Fanuc TP program (LS listing): ConfPr.LS

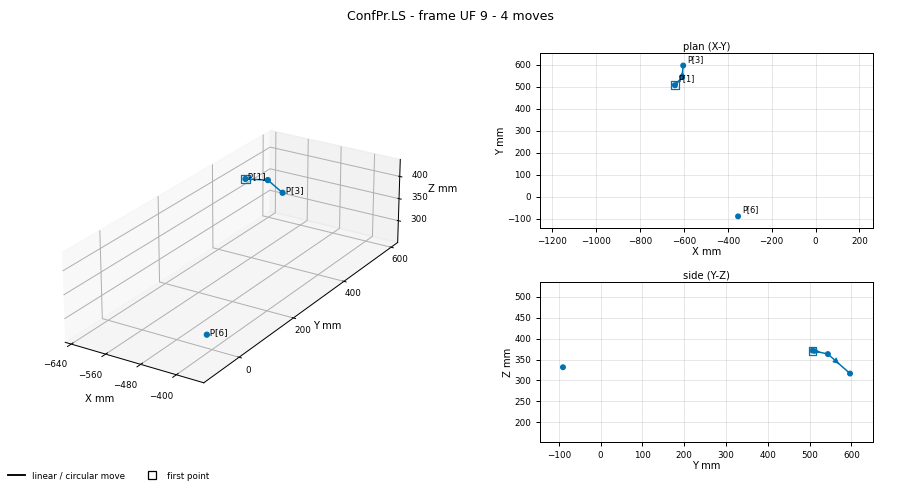
[picture p0: tool path of ConfPr.LS in frame UF 9, 4 of 6 moves have a stored position in this frame; points joined in program order, loops and branches not executed]
/PROG  ConfPr
/ATTR
OWNER		= MNEDITOR;
COMMENT		= "RoboDK sequence";
PROG_SIZE	= 0;
CREATE		= DATE 31-12-14  TIME 12:00:00;
MODIFIED	= DATE 31-12-14  TIME 12:00:00;
FILE_NAME	= ConfPr;
VERSION		= 0;
LINE_COUNT	= 25;
MEMORY_SIZE	= 0;
PROTECT		= READ_WRITE;
TCD:  STACK_SIZE	= 0,
      TASK_PRIORITY	= 50,
      TIME_SLICE	= 0,
      BUSY_LAMP_OFF	= 0,
      ABORT_REQUEST	= 0,
      PAUSE_REQUEST	= 0;
DEFAULT_GROUP	= 1,*,*,*,*;
CONTROL_CODE	= 00000000 00000000;
/MN
   1:  ! Program generated by RoboDK v6.0.7 for Fanuc M-1iA/0.5S on XX ;
   2:  ! /XX/XXXX 18:00:00 ;
   3:  ! Using nominal kinematics. ;
   4:  PR[9,1]=1234.570 ;
   5:  PR[9,2]=-98.765 ;
   6:  PR[9,3]=50.500 ;
   7:  PR[9,4]=0.000 ;
   8:  PR[9,5]=0.000 ;
   9:  PR[9,6]=30.000 ;
  10:  UFRAME[9]=PR[9] ;
  11:  UFRAME_NUM=9 ;
  12:  PR[9,1]=10.000 ;
  13:  PR[9,2]=20.000 ;
  14:  PR[9,3]=150.000 ;
  15:  PR[9,4]=0.000 ;
  16:  PR[9,5]=0.000 ;
  17:  PR[9,6]=0.000 ;
  18:  UTOOL[9]=PR[9] ;
  19:  UTOOL_NUM=9 ;
  20:L P[1] 200mm/sec FINE ;
  21:L P[2] 200mm/sec FINE ;
  22:L P[3] 200mm/sec FINE ;
  23:J P[4] 20% FINE ;
  24:J P[5] 20% FINE ;
  25:C P[6]
       P[7] 200mm/sec FINE ;
/POS
P[1]{
   GP1:
    UF : 9, UT : 9,        CONFIG : 'L, 0, 0, 0',
	X =  -640.584  mm,	Y =   506.980  mm,	Z =   371.534  mm,
	W =  -165.000 deg,	P =    50.000 deg,	R =   150.000 deg
};
P[2]{
   GP1:
    UF : 9, UT : 9,        CONFIG : 'L, 0, 0, 1',
	X =  -607.850  mm,	Y =   543.849  mm,	Z =   363.215  mm,
	W =  -165.000 deg,	P =    50.000 deg,	R =   150.000 deg
};
P[3]{
   GP1:
    UF : 9, UT : 9,        CONFIG : 'R, 0, 0, -1',
	X =  -602.951  mm,	Y =   596.788  mm,	Z =   316.595  mm,
	W =  -165.000 deg,	P =    50.000 deg,	R =   150.000 deg
};
P[4]{
   GP1:
    UF : 9, UT : 9,
	J1=    10.000000 deg,	J2=    20.000000 deg,	J3=    -30.000000  mm,
	J4=    40.000000 deg
};
P[5]{
   GP1:
    UF : 9, UT : 9,
	J1=    -170.000000 deg,	J2=    45.000000 deg,	J3=    -45.000000  mm,
	J4=    -170.000000 deg
};
P[6]{
   GP1:
    UF : 9, UT : 9,        CONFIG : 'R, 0, 0, 1',
	X =  -353.026  mm,	Y =   -90.135  mm,	Z =   331.702  mm,
	W =  -169.444 deg,	P =    40.650 deg,	R =   178.023 deg
};
P[7]{
   GP1:
    UF : 9, UT : 9,        CONFIG : 'L, 0, 0, -1',
	X =  -624.230  mm,	Y =   571.208  mm,	Z =   454.620  mm,
	W =   -82.711 deg,	P =    44.567 deg,	R =  -122.815 deg
};
/END
